(* IEC 61131-3 sources: beedance/examples/simple, 1 file *)

(* ---- my_program.st ---- *)
PROGRAM Main
(* my_program.st *)
VAR
    A : INT := 10;
    B : INT := 20;
END_VAR

A + B;
END_PROGRAM
